// TIA Portal V21 export
// export: Created 2026-11-08T21:35:23.372885Z, ExportSetting WithDefaults, DisplayName Totally Integrated Automation Portal, DisplayVersion V21 Update 3, DisplayName STEP 7 Professional, DisplayVersion V21 Update 3, DisplayName STEP 7 Safety, DisplayVersion V21, DisplayName Tech WebApplication, DisplayVersion V21, DisplayName WinCC Basic/Comfort/Advanced, DisplayVersion V21 Update 3, DisplayName WinCC Unified, DisplayVersion V21 Update 3
FUNCTION_BLOCK "FB_StlC_017"   // FB56, STL
TITLE = STL call IS_NULL
{ S7_Optimized_Access := 'TRUE' }
VERSION : 0.1
// stored: AutoNumber true, IsRetainMemResEnabled false, MemoryReserve 100, UDAEnableTagReadback false
   VAR_INPUT
      "a" : Bool;
      i1 : Int;
      i2 : Int;
      di1 : DInt;
      r1 : Real;
      w1 : Word;
      dw1 : DWord;
      b1 : Byte;
      u1 : UInt;
      ud1 : UDInt;
   END_VAR
   VAR_OUTPUT
      q : Bool;
      io : Int;
      dio : DInt;
      ro : Real;
      wo : Word;
      dwo : DWord;
      bo : Byte;
      udo : UDInt;
   END_VAR
   VAR_IN_OUT
      v : Variant;
      arrs : Array[*] of Int;
      pos : DInt;
   END_VAR
   VAR
      src : Array[0..9] of Int;
      dst : Array[0..9] of Int;
      bits : Array[0..31] of Bool;
      bytes : Array[0..9] of Byte;
      err { S7_SetPoint := 'True'} : ErrorStruct;
      rt : LReal;
      tim { S7_SetPoint := 'True'} : IEC_TIMER;
      words : Array[0..3] of Word;
   END_VAR
BEGIN

NETWORK
TITLE = 017 IS_NULL
      CALL  IS_NULL
      ( OPERAND := #v,
        Ret_Val := #q
      );
END_FUNCTION_BLOCK
